(* IEC 61131-3 sources: Summary-ETFA22/ahorn/test/benchmark/dissertation/PPU/ST (part 7) *)

(* ---- Scenario8_Final_TODO.st ---- *)
FUNCTION_BLOCK Crane

    VAR_OUTPUT
        AnalogCranePressure : INT := INT#0;
        CraneLower : BOOL := FALSE;
        CraneTurnClockwise : BOOL := FALSE;
        CraneTurnCounterclockwise : BOOL := FALSE;
        MagazinVacuumOff : BOOL := FALSE;
        MagazinVacuumOn : BOOL := FALSE;
        StartCommandCrane : BOOL := FALSE;
    END_VAR

    VAR_INPUT
        CraneDown : BOOL := FALSE;
        CraneOnConveyor : BOOL := FALSE;
        CraneOnMagazin : BOOL := FALSE;
        CranePositionStamp : BOOL := FALSE;
        CraneSucked : BOOL := FALSE;
        CraneUp : BOOL := FALSE;
        MagazinCapacitiveSensor : BOOL := FALSE;
        MagazinOpticalSensor : BOOL := FALSE;
        SFCReset : BOOL := FALSE;
        SliderMovedOut : BOOL := FALSE;
        SliderNotMovedOut : BOOL := FALSE;
        StampLowered : BOOL := FALSE;
        StampSliderFilled : BOOL := FALSE;
        StampSliderSensorMovedOut : BOOL := FALSE;
        StartButtonMagazin : BOOL := FALSE;
        StartVar : BOOL := FALSE;
        WorkpieceReady : BOOL := FALSE;
    END_VAR

    VAR
        Duration1 : TIME := TIME#1500.0ms;
        SFCInit : BOOL := FALSE;
        TimeDelay_Timer : TON := (Q:=FALSE, PT:=UINT#0, IN:=FALSE, ET:=UINT#0);
        TimeDelay_Timer_Duration : TIME := TIME#50.0ms;
        TimeDelay_Timer_interconnect : BOOL := FALSE;
        Timer1 : TON := (Q:=FALSE, PT:=UINT#0, IN:=FALSE, ET:=UINT#0);
        actualtime1 : TIME := TIME#;
        interconnect : BOOL := FALSE;
        interconnectCraneStartCommand : BOOL := FALSE;
    END_VAR

    VAR
        SFCPause : BOOL := FALSE;
    END_VAR

    VAR
        __transit : BOOL := FALSE;
        _state : STATES_CRANE := STATES_CRANE#INIT;
    END_VAR

    ACTION Turn_Right_active
        CraneTurnClockwise := TRUE;
        CraneTurnCounterclockwise := FALSE;
    END_ACTION
    ACTION Crane_Turn_Left_White_active
        CraneTurnCounterclockwise := TRUE;
        CraneTurnClockwise := FALSE;
    END_ACTION
    ACTION Crane_Turn_Left_Metallic_active
        CraneTurnCounterclockwise := TRUE;
        CraneTurnClockwise := FALSE;
    END_ACTION
    ACTION Crane_Lift_Conveyor2_active
        CraneLower := FALSE;
    END_ACTION
    ACTION Crane_Turn_Right_From_Stamp_active
        CraneTurnClockwise := TRUE;
        CraneTurnCounterclockwise := FALSE;
    END_ACTION
    ACTION Suck_At_Stamp_active
        MagazinVacuumOn := TRUE;
        MagazinVacuumOff := FALSE;
    END_ACTION
    ACTION CraneTurnLeft_active
        CraneTurnCounterclockwise := TRUE;
        CraneTurnClockwise := FALSE;
    END_ACTION
    ACTION Crane_Turn_Left_From_Stamp_active
        CraneTurnClockwise := TRUE;
        CraneTurnCounterclockwise := FALSE;
    END_ACTION
    ACTION release_Black_active
        MagazinVacuumOn := FALSE;
        MagazinVacuumOff := TRUE;
    END_ACTION
    ACTION Crane_On_Stamp_Stop_Black_active
        CraneTurnClockwise := FALSE;
        CraneTurnCounterclockwise := FALSE;
    END_ACTION
    ACTION Reset_interconnect_active
        interconnect := FALSE;
        Timer1(IN := FALSE, PT := TIME#1ms);
    END_ACTION
    ACTION Crane_On_Stamp_White_active
        CraneTurnCounterclockwise := FALSE;
        CraneTurnClockwise := FALSE;
        CraneLower := TRUE;
    END_ACTION
    ACTION Crane_On_Stamp_Metallic_active
        CraneTurnCounterclockwise := FALSE;
        CraneTurnClockwise := FALSE;
        CraneLower := TRUE;
    END_ACTION
    ACTION Crane_Lift_Magazin_Metallic_active_0
        CraneLower := FALSE;
    END_ACTION
    ACTION TimeDelay_active
        TimeDelay_Timer(IN := TRUE, PT := TimeDelay_Timer_Duration);
        TimeDelay_Timer_interconnect := TimeDelay_Timer.Q;
    END_ACTION
    ACTION CraneLiftConveyor_active
        CraneLower := FALSE;
    END_ACTION
    ACTION Crane_Turn_Left_Back_To_Stamp_active
        CraneTurnCounterclockwise := TRUE;
        CraneTurnClockwise := FALSE;
    END_ACTION
    ACTION Crane_Init_2_active
        CraneLower := FALSE;
    END_ACTION
    ACTION Crane_Lower_active
        MagazinVacuumOn := TRUE;
        MagazinVacuumOff := FALSE;
        CraneLower := TRUE;
        AnalogCranePressure := INT#0;
    END_ACTION
    ACTION Crane_Lift_At_Stamp2_active
        CraneLower := FALSE;
    END_ACTION
    ACTION Crane_On_Stamp_Metallic2_active
        CraneTurnCounterclockwise := FALSE;
        CraneTurnClockwise := FALSE;
    END_ACTION
    ACTION CraneLiftMagazin_active
        CraneLower := FALSE;
    END_ACTION
    ACTION release_active
        MagazinVacuumOff := TRUE;
        MagazinVacuumOn := FALSE;
    END_ACTION
    ACTION Lower_Crane_active
        CraneLower := TRUE;
    END_ACTION
    ACTION Start_Crane_active
        CraneLower := FALSE;
        MagazinVacuumOff := TRUE;
        MagazinVacuumOn := FALSE;
        CraneTurnCounterclockwise := FALSE;
        CraneTurnClockwise := FALSE;
        StartVar := FALSE;
        StartCommandCrane := FALSE;
        IF (StartButtonMagazin = TRUE) THEN
            interconnectCraneStartCommand := TRUE;
        END_IF
    END_ACTION
    ACTION Crane_Go_Up_White_active
        CraneLower := FALSE;
    END_ACTION
    ACTION Crane_Init_active
        CraneLower := TRUE;
        interconnectCraneStartCommand := FALSE;
        AnalogCranePressure := INT#6000;
    END_ACTION
    ACTION Crane_Turn_Left_NOT_Metallic_Black_active
        CraneTurnCounterclockwise := TRUE;
        CraneTurnClockwise := FALSE;
    END_ACTION
    ACTION release_Workpiece_White_active
        MagazinVacuumOff := TRUE;
        MagazinVacuumOn := FALSE;
    END_ACTION
    ACTION Crane_On_Stamp_Metallic2_Lower_active
        CraneLower := TRUE;
    END_ACTION
    ACTION Crane_Turn_Left_Metallic2_active
        CraneTurnCounterclockwise := TRUE;
        CraneTurnClockwise := FALSE;
    END_ACTION
    ACTION Crane_Lift_NOT_Metallic_Black_active
        CraneLower := FALSE;
    END_ACTION
    ACTION Magazin_Stop_active
        CraneTurnClockwise := FALSE;
        CraneTurnCounterClockwise := FALSE;
    END_ACTION
    ACTION Crane_On_Conveyor_Not_Metallica_Black_active
        CraneTurnCounterclockwise := FALSE;
        CraneTurnClockwise := FALSE;
        CraneLower := TRUE;
    END_ACTION
    ACTION release_Workpiece_active
        MagazinVacuumOff := TRUE;
        MagazinVacuumOn := FALSE;
    END_ACTION
    ACTION No_Workpiece_ready_active_0
        MagazinVacuumOn := FALSE;
        MagazinVacuumOff := FALSE;
        CraneLower := FALSE;
    END_ACTION
    ACTION CraneOnConveyor_active
        CraneTurnCounterclockwise := FALSE;
        CraneTurnClockwise := FALSE;
        CraneLower := TRUE;
    END_ACTION
    ACTION Crane_Go_Up_active
        CraneLower := FALSE;
    END_ACTION
    ACTION Turn_Right_Final_active
        CraneTurnClockwise := TRUE;
        CraneTurnCounterclockwise := FALSE;
        AnalogCranePressure := INT#0;
    END_ACTION
    ACTION Suck_At_Stamp2_active
        MagazinVacuumOn := TRUE;
        MagazinVacuumOff := FALSE;
    END_ACTION
    ACTION Stamp_Pressure_Profile_Set_White_active
        AnalogCranePressure := INT#6000;
    END_ACTION
    ACTION Interstep_active
        StartCommandCrane := TRUE;
    END_ACTION
    ACTION Turn_Right_Black_active
        CraneTurnClockwise := TRUE;
        CraneTurnCounterclockwise := FALSE;
    END_ACTION
    ACTION Crane_On_Conveyor_Metallic2_active
        CraneTurnCounterclockwise := FALSE;
        CraneTurnClockwise := FALSE;
        CraneLower := TRUE;
    END_ACTION
    ACTION Crane_Lift_Conveyor_Black_active
        CraneLower := FALSE;
    END_ACTION
    ACTION Magazin_Stop_Final_active
        CraneTurnClockwise := FALSE;
        CraneTurnCounterClockwise := FALSE;
    END_ACTION
    ACTION Stamp_Pressure_Profile_Set_Metallic_active
        AnalogCranePressure := INT#7000;
    END_ACTION
    ACTION Crane_Lift_At_Stamp_active
        CraneLower := FALSE;
    END_ACTION
    ACTION Magazin_Stop_Black_active
        CraneTurnClockwise := FALSE;
        CraneTurnCounterclockwise := FALSE;
        MagazinVacuumOn := TRUE;
        MagazinVacuumOff := FALSE;
        CraneLower := TRUE;
    END_ACTION
    ACTION Crane_Lift_Magazin_White_active
        CraneLower := FALSE;
    END_ACTION
    ACTION pause_active
        Timer1(IN := CraneUP, PT := Duration1);
        interconnect := Timer1.Q;
    END_ACTION
    ACTION Crane_On_Conveyor_Metallic_active_0
        CraneTurnCounterclockwise := FALSE;
        CraneTurnClockwise := FALSE;
        CraneLower := TRUE;
    END_ACTION
    ACTION release2_active
        MagazinVacuumOff := TRUE;
        MagazinVacuumOn := FALSE;
    END_ACTION
    IF (SFCInit OR SFCReset) THEN
        AnalogCranePressure := INT#0;
        CraneDown := FALSE;
        CraneLower := FALSE;
        CraneOnConveyor := FALSE;
        CraneOnMagazin := FALSE;
        CranePositionStamp := FALSE;
        CraneSucked := FALSE;
        CraneTurnClockwise := FALSE;
        CraneTurnCounterclockwise := FALSE;
        CraneUp := FALSE;
        Duration1 := TIME#1500ms;
        MagazinCapacitiveSensor := FALSE;
        MagazinOpticalSensor := FALSE;
        MagazinVacuumOff := FALSE;
        MagazinVacuumOn := FALSE;
        SFCInit := FALSE;
        SFCReset := FALSE;
        SliderMovedOut := FALSE;
        SliderNotMovedOut := FALSE;
        StampLowered := FALSE;
        StampSliderFilled := FALSE;
        StampSliderSensorMovedOut := FALSE;
        StartButtonMagazin := FALSE;
        StartCommandCrane := FALSE;
        StartVar := FALSE;
        TimeDelay_Timer.ET := UINT#0;
        TimeDelay_Timer.IN := FALSE;
        TimeDelay_Timer.PT := UINT#0;
        TimeDelay_Timer.Q := FALSE;
        TimeDelay_Timer_Duration := TIME#50ms;
        TimeDelay_Timer_interconnect := FALSE;
        Timer1.ET := UINT#0;
        Timer1.IN := FALSE;
        Timer1.PT := UINT#0;
        Timer1.Q := FALSE;
        WorkpieceReady := FALSE;
        __transit := FALSE;
        _state := STATES_CRANE#INIT;
        actualtime1 := TIME#0ms;
        interconnect := FALSE;
        interconnectCraneStartCommand := FALSE;
    END_IF
    IF NOT (SFCInit OR SFCPause) THEN
        //Running pipeline step: edu.kit.iti.formal.automation.st.IntroduceStateEnumVariable

        //End of: edu.kit.iti.formal.automation.st.IntroduceStateEnumVariable

        //Running pipeline step: edu.kit.iti.formal.automation.st.TranslationSfcToStOld$IntroduceTransitVariable

        //End of: edu.kit.iti.formal.automation.st.TranslationSfcToStOld$IntroduceTransitVariable

        //Running pipeline step: edu.kit.iti.formal.automation.st.TranslationSfcToStOld$TheBigStateCase

        CASE _state OF
            STATES_CRANE#Init:
                __transit := FALSE;
                IF TRUE THEN
                    __transit := TRUE;
                    _state := STATES_CRANE#Start_Crane;
                END_IF

            STATES_CRANE#Start_Crane:
                __transit := FALSE;
                Start_Crane_active();
                IF interconnectCraneStartCommand THEN
                    __transit := TRUE;
                    _state := STATES_CRANE#Crane_Init;
                END_IF

            STATES_CRANE#Crane_Init:
                __transit := FALSE;
                Crane_Init_active();
                IF CraneDown THEN
                    __transit := TRUE;
                    _state := STATES_CRANE#Crane_Init_2;
                END_IF

            STATES_CRANE#Crane_Init_2:
                __transit := FALSE;
                Crane_Init_2_active();
                IF CraneUp THEN
                    __transit := TRUE;
                    _state := STATES_CRANE#Interstep;
                END_IF

            STATES_CRANE#Interstep:
                __transit := FALSE;
                Interstep_active();
                IF StartVar THEN
                    __transit := TRUE;
                    _state := STATES_CRANE#Interstep_2;
                END_IF

            STATES_CRANE#Interstep_2:
                __transit := FALSE;
                IF SliderMovedOut THEN
                    __transit := TRUE;
                    _state := STATES_CRANE#TimeDelay;
                END_IF

            STATES_CRANE#TimeDelay:
                __transit := FALSE;
                TimeDelay_active();
                IF TimeDelay_Timer_interconnect THEN
                    __transit := TRUE;
                    _state := STATES_CRANE#Interstep_3;
                END_IF

            STATES_CRANE#Interstep_3:
                __transit := FALSE;
                IF WorkpieceReady THEN
                    __transit := TRUE;
                    _state := STATES_CRANE#Turn_Right;
                ELSIF NOT WorkpieceReady THEN
                    __transit := TRUE;
                    _state := STATES_CRANE#No_Workpiece_ready;
                END_IF

            STATES_CRANE#Turn_Right:
                __transit := FALSE;
                Turn_Right_active();
                IF CraneOnMagazin THEN
                    __transit := TRUE;
                    _state := STATES_CRANE#Magazin_Stop;
                END_IF

            STATES_CRANE#Magazin_Stop:
                __transit := FALSE;
                Magazin_Stop_active();
                IF TRUE THEN
                    __transit := TRUE;
                    _state := STATES_CRANE#Crane_Lower;
                END_IF

            STATES_CRANE#Crane_Lower:
                __transit := FALSE;
                Crane_Lower_active();
                IF CraneSucked THEN
                    __transit := TRUE;
                    _state := STATES_CRANE#Step0;
                END_IF

            STATES_CRANE#Step0:
                __transit := FALSE;
                IF (NOT MagazinCapacitiveSensor AND NOT MagazinOpticalSensor) THEN
                    __transit := TRUE;
                    _state := STATES_CRANE#Crane_Lift_Magazin;
                ELSIF (MagazinCapacitiveSensor AND MagazinOpticalSensor) THEN
                    __transit := TRUE;
                    _state := STATES_CRANE#Stamp_Pressure_Profile_Set_Metallic;
                ELSIF (NOT MagazinCapacitiveSensor AND MagazinOpticalSensor) THEN
                    __transit := TRUE;
                    _state := STATES_CRANE#Stamp_Pressure_Profile_Set_White;
                ELSIF (MagazinCapacitiveSensor AND MagazinOpticalSensor) THEN
                    __transit := TRUE;
                    _state := STATES_CRANE#Stamp_Pressure_Profile_Set_Metallic;
                ELSIF (NOT MagazinCapacitiveSensor AND MagazinOpticalSensor) THEN
                    __transit := TRUE;
                    _state := STATES_CRANE#Stamp_Pressure_Profile_Set_White;
                END_IF

            STATES_CRANE#Crane_Lift_Magazin:
                __transit := FALSE;
                CraneLiftMagazin_active();
                IF CraneUp THEN
                    __transit := TRUE;
                    _state := STATES_CRANE#Crane_Turn_Left_NOT_Metallic;
                END_IF

            STATES_CRANE#Crane_Turn_Left_NOT_Metallic:
                __transit := FALSE;
                CraneTurnLeft_active();
                IF CraneOnConveyor THEN
                    __transit := TRUE;
                    _state := STATES_CRANE#Crane_On_Conveyor;
                END_IF

            STATES_CRANE#Crane_On_Conveyor:
                __transit := FALSE;
                CraneOnConveyor_active();
                IF CraneDown THEN
                    __transit := TRUE;
                    _state := STATES_CRANE#release;
                END_IF

            STATES_CRANE#Stamp_Pressure_Profile_Set_Metallic:
                __transit := FALSE;
                Stamp_Pressure_Profile_Set_Metallic_active();
                IF TRUE THEN
                    __transit := TRUE;
                    _state := STATES_CRANE#Crane_Lift_Magazin_Metallic;
                END_IF

            STATES_CRANE#Crane_Lift_Magazin_Metallic:
                __transit := FALSE;
                Crane_Lift_Magazin_Metallic_active_0();
                IF CraneUp THEN
                    __transit := TRUE;
                    _state := STATES_CRANE#Crane_Turn_Left_Metallic;
                END_IF

            STATES_CRANE#Crane_Turn_Left_Metallic:
                __transit := FALSE;
                Crane_Turn_Left_Metallic_active();
                IF CranePositionStamp THEN
                    __transit := TRUE;
                    _state := STATES_CRANE#Crane_On_Stamp_Metallic;
                END_IF

            STATES_CRANE#Crane_On_Stamp_Metallic:
                __transit := FALSE;
                Crane_On_Stamp_Metallic_active();
                IF CraneDown THEN
                    __transit := TRUE;
                    _state := STATES_CRANE#release_Workpiece;
                END_IF

            STATES_CRANE#release_Workpiece:
                __transit := FALSE;
                release_Workpiece_active();
                IF TRUE THEN
                    __transit := TRUE;
                    _state := STATES_CRANE#Crane_Go_Up;
                END_IF

            STATES_CRANE#Crane_Go_Up:
                __transit := FALSE;
                Crane_Go_Up_active();
                IF CraneUp THEN
                    __transit := TRUE;
                    _state := STATES_CRANE#Step3;
                END_IF

            STATES_CRANE#Stamp_Pressure_Profile_Set_White:
                __transit := FALSE;
                Stamp_Pressure_Profile_Set_White_active();
                IF TRUE THEN
                    __transit := TRUE;
                    _state := STATES_CRANE#Crane_Lift_Magazine_White;
                END_IF

            STATES_CRANE#Crane_Lift_Magazine_White:
                __transit := FALSE;
                Crane_Lift_Magazin_White_active();
                IF CraneUp THEN
                    __transit := TRUE;
                    _state := STATES_CRANE#Crane_Turn_Left_White;
                END_IF

            STATES_CRANE#Crane_Turn_Left_White:
                __transit := FALSE;
                Crane_Turn_Left_White_active();
                IF CranePositionStamp THEN
                    __transit := TRUE;
                    _state := STATES_CRANE#Crane_On_Stamp_White;
                END_IF

            STATES_CRANE#Crane_On_Stamp_White:
                __transit := FALSE;
                Crane_On_Stamp_White_active();
                IF CraneDown THEN
                    __transit := TRUE;
                    _state := STATES_CRANE#release_Workpiece_White;
                END_IF

            STATES_CRANE#release_Workpiece_White:
                __transit := FALSE;
                release_Workpiece_White_active();
                IF TRUE THEN
                    __transit := TRUE;
                    _state := STATES_CRANE#Crane_Go_Up_White;
                END_IF

            STATES_CRANE#Crane_Go_Up_White:
                __transit := FALSE;
                Crane_Go_Up_White_active();
                IF CraneUp THEN
                    __transit := TRUE;
                    _state := STATES_CRANE#Step3;
                END_IF

            STATES_CRANE#Step3:
                __transit := FALSE;
                IF WorkpieceReady THEN
                    __transit := TRUE;
                    _state := STATES_CRANE#Step2;
                ELSIF NOT WorkpieceReady THEN
                    __transit := TRUE;
                    _state := STATES_CRANE#Step4;
                END_IF

            STATES_CRANE#Step2:
                __transit := FALSE;
                IF (MagazinCapacitiveSensor OR MagazinOpticalSensor) THEN
                    __transit := TRUE;
                    _state := STATES_CRANE#pause;
                ELSIF (NOT MagazinCapacitiveSensor AND NOT MagazinOpticalSensor) THEN
                    __transit := TRUE;
                    _state := STATES_CRANE#Turn_Right_Black;
                END_IF

            STATES_CRANE#pause:
                __transit := FALSE;
                pause_active();
                IF interconnect THEN
                    __transit := TRUE;
                    _state := STATES_CRANE#Reset_interconnect;
                ELSIF interconnect THEN
                    __transit := TRUE;
                    _state := STATES_CRANE#Reset_interconnect;
                END_IF

            STATES_CRANE#Turn_Right_Black:
                __transit := FALSE;
                Turn_Right_Black_active();
                IF CraneOnMagazin THEN
                    __transit := TRUE;
                    _state := STATES_CRANE#Magazin_Stop_Black;
                END_IF

            STATES_CRANE#Magazin_Stop_Black:
                __transit := FALSE;
                Magazin_Stop_Black_active();
                IF CraneSucked THEN
                    __transit := TRUE;
                    _state := STATES_CRANE#Crane_Lift_NOT_Metallic_Black;
                END_IF

            STATES_CRANE#Crane_Lift_NOT_Metallic_Black:
                __transit := FALSE;
                Crane_Lift_NOT_Metallic_Black_active();
                IF CraneUp THEN
                    __transit := TRUE;
                    _state := STATES_CRANE#Crane_Turn_Left_NOT_Metallic_Black;
                END_IF

            STATES_CRANE#Crane_Turn_Left_NOT_Metallic_Black:
                __transit := FALSE;
                Crane_Turn_Left_NOT_Metallic_Black_active();
                IF CraneOnConveyor THEN
                    __transit := TRUE;
                    _state := STATES_CRANE#Crane_On_Conveyor_Not_Metallica_Black;
                END_IF

            STATES_CRANE#Crane_On_Conveyor_Not_Metallica_Black:
                __transit := FALSE;
                Crane_On_Conveyor_Not_Metallica_Black_active();
                IF CraneDown THEN
                    __transit := TRUE;
                    _state := STATES_CRANE#release_Black;
                END_IF

            STATES_CRANE#release_Black:
                __transit := FALSE;
                release_Black_active();
                IF TRUE THEN
                    __transit := TRUE;
                    _state := STATES_CRANE#Crane_Lift_Conveyor_Black;
                END_IF

            STATES_CRANE#Crane_Lift_Conveyor_Black:
                __transit := FALSE;
                Crane_Lift_Conveyor_Black_active();
                IF CraneUp THEN
                    __transit := TRUE;
                    _state := STATES_CRANE#Crane_Turn_Left_Back_To_Stamp;
                END_IF

            STATES_CRANE#Crane_Turn_Left_Back_To_Stamp:
                __transit := FALSE;
                Crane_Turn_Left_Back_To_Stamp_active();
                IF CranePositionStamp THEN
                    __transit := TRUE;
                    _state := STATES_CRANE#Crane_On_Stamp_Stop_Black;
                END_IF

            STATES_CRANE#Crane_On_Stamp_Stop_Black:
                __transit := FALSE;
                Crane_On_Stamp_Stop_Black_active();
                IF TRUE THEN
                    __transit := TRUE;
                    _state := STATES_CRANE#Reset_interconnect;
                ELSIF TRUE THEN
                    __transit := TRUE;
                    _state := STATES_CRANE#Reset_interconnect;
                END_IF

            STATES_CRANE#Step4:
                __transit := FALSE;
                IF TRUE THEN
                    __transit := TRUE;
                    _state := STATES_CRANE#Interstep;
                END_IF

            STATES_CRANE#Reset_interconnect:
                __transit := FALSE;
                Reset_interconnect_active();
                IF SliderMovedOut THEN
                    __transit := TRUE;
                    _state := STATES_CRANE#Lower_Crane;
                END_IF

            STATES_CRANE#Lower_Crane:
                __transit := FALSE;
                Lower_Crane_active();
                IF CraneDown THEN
                    __transit := TRUE;
                    _state := STATES_CRANE#Suck_At_Stamp;
                END_IF

            STATES_CRANE#Suck_At_Stamp:
                __transit := FALSE;
                Suck_At_Stamp_active();
                IF CraneSucked THEN
                    __transit := TRUE;
                    _state := STATES_CRANE#Crane_Lift_At_Stamp;
                END_IF

            STATES_CRANE#Crane_Lift_At_Stamp:
                __transit := FALSE;
                Crane_Lift_At_Stamp_active();
                IF CraneUp THEN
                    __transit := TRUE;
                    _state := STATES_CRANE#Crane_Turn_Left_From_Stamp;
                END_IF

            STATES_CRANE#Crane_Turn_Left_From_Stamp:
                __transit := FALSE;
                Crane_Turn_Left_From_Stamp_active();
                IF CraneOnConveyor THEN
                    __transit := TRUE;
                    _state := STATES_CRANE#Crane_On_Conveyor_Metallic;
                END_IF

            STATES_CRANE#Crane_On_Conveyor_Metallic:
                __transit := FALSE;
                Crane_On_Conveyor_Metallic_active_0();
                IF CraneDown THEN
                    __transit := TRUE;
                    _state := STATES_CRANE#release;
                END_IF

            STATES_CRANE#release:
                __transit := FALSE;
                release_active();
                IF TRUE THEN
                    __transit := TRUE;
                    _state := STATES_CRANE#Crane_Lift_Conveyor;
                END_IF

            STATES_CRANE#Crane_Lift_Conveyor:
                __transit := FALSE;
                CraneLiftConveyor_active();
                IF TRUE THEN
                    __transit := TRUE;
                    _state := STATES_CRANE#Interstep;
                END_IF

            STATES_CRANE#No_Workpiece_ready:
                __transit := FALSE;
                No_Workpiece_ready_active_0();
                IF StampSliderFilled THEN
                    __transit := TRUE;
                    _state := STATES_CRANE#Crane_Turn_Left_Metallic2;
                ELSIF NOT StampSliderFilled THEN
                    __transit := TRUE;
                    _state := STATES_CRANE#Turn_Right_Final;
                END_IF

            STATES_CRANE#Crane_Turn_Left_Metallic2:
                __transit := FALSE;
                Crane_Turn_Left_Metallic2_active();
                IF CranePositionStamp THEN
                    __transit := TRUE;
                    _state := STATES_CRANE#Crane_On_Stamp_Metallic2;
                END_IF

            STATES_CRANE#Crane_On_Stamp_Metallic2:
                __transit := FALSE;
                Crane_On_Stamp_Metallic2_active();
                IF StampLowered THEN
                    __transit := TRUE;
                    _state := STATES_CRANE#Interstep_4;
                END_IF

            STATES_CRANE#Interstep_4:
                __transit := FALSE;
                IF StampSliderSensorMovedOut THEN
                    __transit := TRUE;
                    _state := STATES_CRANE#Crane_On_Stamp_Metallic2_Lower;
                END_IF

            STATES_CRANE#Crane_On_Stamp_Metallic2_Lower:
                __transit := FALSE;
                Crane_On_Stamp_Metallic2_Lower_active();
                IF CraneDown THEN
                    __transit := TRUE;
                    _state := STATES_CRANE#Suck_At_Stamp2;
                END_IF

            STATES_CRANE#Suck_At_Stamp2:
                __transit := FALSE;
                Suck_At_Stamp2_active();
                IF CraneSucked THEN
                    __transit := TRUE;
                    _state := STATES_CRANE#Crane_Lift_At_Stamp2;
                END_IF

            STATES_CRANE#Crane_Lift_At_Stamp2:
                __transit := FALSE;
                Crane_Lift_At_Stamp2_active();
                IF CraneUp THEN
                    __transit := TRUE;
                    _state := STATES_CRANE#Crane_Turn_Right_From_Stamp;
                END_IF

            STATES_CRANE#Crane_Turn_Right_From_Stamp:
                __transit := FALSE;
                Crane_Turn_Right_From_Stamp_active();
                IF CraneOnConveyor THEN
                    __transit := TRUE;
                    _state := STATES_CRANE#Crane_On_Conveyor_Metallic2;
                END_IF

            STATES_CRANE#Crane_On_Conveyor_Metallic2:
                __transit := FALSE;
                Crane_On_Conveyor_Metallic2_active();
                IF CraneDown THEN
                    __transit := TRUE;
                    _state := STATES_CRANE#release2;
                END_IF

            STATES_CRANE#release2:
                __transit := FALSE;
                release2_active();
                IF TRUE THEN
                    __transit := TRUE;
                    _state := STATES_CRANE#Crane_Lift_Conveyor2;
                END_IF

            STATES_CRANE#Crane_Lift_Conveyor2:
                __transit := FALSE;
                Crane_Lift_Conveyor2_active();
                IF TRUE THEN
                    __transit := TRUE;
                    _state := STATES_CRANE#Interstep;
                ELSIF TRUE THEN
                    __transit := TRUE;
                    _state := STATES_CRANE#Interstep;
                END_IF

            STATES_CRANE#Turn_Right_Final:
                __transit := FALSE;
                Turn_Right_Final_active();
                IF CraneOnMagazin THEN
                    __transit := TRUE;
                    _state := STATES_CRANE#Magazin_Stop_Final;
                END_IF

            STATES_CRANE#Magazin_Stop_Final:
                __transit := FALSE;
                Magazin_Stop_Final_active();
                IF TRUE THEN
                    __transit := TRUE;
                    _state := STATES_CRANE#Start_Crane;
                END_IF

                    END_CASE
        //End of: edu.kit.iti.formal.automation.st.TranslationSfcToStOld$TheBigStateCase

        //Running pipeline step: edu.kit.iti.formal.automation.st.SfcFlagIntroduction

    END_IF
    //End of: edu.kit.iti.formal.automation.st.SfcFlagIntroduction

END_FUNCTION_BLOCK

FUNCTION_BLOCK Magazin

    VAR_INPUT
        CraneDown : BOOL := FALSE;
        CraneOnConveyor : BOOL := FALSE;
        CraneOnMagazin : BOOL := FALSE;
        CraneSucked : BOOL := FALSE;
        CraneUp : BOOL := FALSE;
        SFCReset : BOOL := FALSE;
        SliderMovedOut : BOOL := FALSE;
        SliderNotMovedOut : BOOL := FALSE;
        StartButtonMagazin : BOOL := FALSE;
        StartVar : BOOL := FALSE;
        WorkpieceReady : BOOL := FALSE;
    END_VAR

    VAR_OUTPUT
        CraneLower : BOOL := FALSE;
        CraneTurnClockwise : BOOL := FALSE;
        CraneTurnCounterclockwise : BOOL := FALSE;
        MagazinGreenLamp : BOOL := FALSE;
        MagazinSlider : BOOL := FALSE;
        MagazinVacuumOff : BOOL := FALSE;
        MagazinVacuumOn : BOOL := FALSE;
        MagazinWhiteLamp : BOOL := FALSE;
        StartCommandMagazin : BOOL := FALSE;
    END_VAR

    VAR
        SFCInit : BOOL := FALSE;
        interconnectMagazinStartCommand : BOOL := FALSE;
    END_VAR

    VAR
        SFCPause : BOOL := FALSE;
    END_VAR

    VAR
        __transit : BOOL := FALSE;
        _state : STATES_MAGAZIN := STATES_MAGAZIN#INIT;
    END_VAR

    ACTION Magazin_Init_2_active
        MagazinSlider := FALSE;
    END_ACTION
    ACTION Start_Magazin_active
        MagazinSlider := FALSE;
        MagazinGreenLamp := FALSE;
        StartVar := FALSE;
        StartCommandMagazin := FALSE;
        IF (StartButtonMagazin = TRUE) THEN
            interconnectMagazinStartCommand := TRUE;
        END_IF
    END_ACTION
    ACTION Green_Lamp_active
        MagazinGreenLamp := TRUE;
        interconnectMagazinStartCommand := FALSE;
    END_ACTION
    ACTION SliderMoveBack_active
        IF ((SliderMovedOut = TRUE) AND (SliderNotMovedOut = FALSE)) THEN
            MagazinSlider := FALSE;
        END_IF
    END_ACTION
    ACTION convey_active
        IF SliderNotMovedOut THEN
            MagazinSlider := TRUE;
        END_IF
    END_ACTION
    ACTION Magazin_Init_active
        MagazinSlider := TRUE;
    END_ACTION
    ACTION Interstep_active
        StartCommandMagazin := TRUE;
    END_ACTION
    IF (SFCInit OR SFCReset) THEN
        CraneDown := FALSE;
        CraneLower := FALSE;
        CraneOnConveyor := FALSE;
        CraneOnMagazin := FALSE;
        CraneSucked := FALSE;
        CraneTurnClockwise := FALSE;
        CraneTurnCounterclockwise := FALSE;
        CraneUp := FALSE;
        MagazinGreenLamp := FALSE;
        MagazinSlider := FALSE;
        MagazinVacuumOff := FALSE;
        MagazinVacuumOn := FALSE;
        MagazinWhiteLamp := FALSE;
        SFCInit := FALSE;
        SFCReset := FALSE;
        SliderMovedOut := FALSE;
        SliderNotMovedOut := FALSE;
        StartButtonMagazin := FALSE;
        StartCommandMagazin := FALSE;
        StartVar := FALSE;
        WorkpieceReady := FALSE;
        __transit := FALSE;
        _state := STATES_MAGAZIN#INIT;
        interconnectMagazinStartCommand := FALSE;
    END_IF
    IF NOT (SFCInit OR SFCPause) THEN
        //Running pipeline step: edu.kit.iti.formal.automation.st.IntroduceStateEnumVariable

        //End of: edu.kit.iti.formal.automation.st.IntroduceStateEnumVariable

        //Running pipeline step: edu.kit.iti.formal.automation.st.TranslationSfcToStOld$IntroduceTransitVariable

        //End of: edu.kit.iti.formal.automation.st.TranslationSfcToStOld$IntroduceTransitVariable

        //Running pipeline step: edu.kit.iti.formal.automation.st.TranslationSfcToStOld$TheBigStateCase

        CASE _state OF
            STATES_MAGAZIN#Init:
                __transit := FALSE;
                IF TRUE THEN
                    __transit := TRUE;
                    _state := STATES_MAGAZIN#Start_Magazin;
                END_IF

            STATES_MAGAZIN#Start_Magazin:
                __transit := FALSE;
                Start_Magazin_active();
                IF interconnectMagazinStartCommand THEN
                    __transit := TRUE;
                    _state := STATES_MAGAZIN#Green_Lamp;
                END_IF

            STATES_MAGAZIN#Green_Lamp:
                __transit := FALSE;
                Green_Lamp_active();
                IF TRUE THEN
                    __transit := TRUE;
                    _state := STATES_MAGAZIN#Magazin_Init;
                END_IF

            STATES_MAGAZIN#Magazin_Init:
                __transit := FALSE;
                Magazin_Init_active();
                IF TRUE THEN
                    __transit := TRUE;
                    _state := STATES_MAGAZIN#Magazin_Init_2;
                END_IF

            STATES_MAGAZIN#Magazin_Init_2:
                __transit := FALSE;
                Magazin_Init_2_active();
                IF TRUE THEN
                    __transit := TRUE;
                    _state := STATES_MAGAZIN#Interstep;
                END_IF

            STATES_MAGAZIN#Interstep:
                __transit := FALSE;
                Interstep_active();
                IF StartVar THEN
                    __transit := TRUE;
                    _state := STATES_MAGAZIN#convey;
                END_IF

            STATES_MAGAZIN#convey:
                __transit := FALSE;
                convey_active();
                IF CraneOnMagazin THEN
                    __transit := TRUE;
                    _state := STATES_MAGAZIN#Step0;
                END_IF

            STATES_MAGAZIN#Step0:
                __transit := FALSE;
                IF CraneDown THEN
                    __transit := TRUE;
                    _state := STATES_MAGAZIN#Slider_Move_Back;
                END_IF

            STATES_MAGAZIN#Slider_Move_Back:
                __transit := FALSE;
                SliderMoveBack_active();
                IF CraneUp THEN
                    __transit := TRUE;
                    _state := STATES_MAGAZIN#Step1;
                END_IF

            STATES_MAGAZIN#Step1:
                __transit := FALSE;
                IF CraneOnConveyor THEN
                    __transit := TRUE;
                    _state := STATES_MAGAZIN#Interstep;
                END_IF

                    END_CASE
        //End of: edu.kit.iti.formal.automation.st.TranslationSfcToStOld$TheBigStateCase

        //Running pipeline step: edu.kit.iti.formal.automation.st.SfcFlagIntroduction

    END_IF
    //End of: edu.kit.iti.formal.automation.st.SfcFlagIntroduction

END_FUNCTION_BLOCK

FUNCTION_BLOCK Stamp

    VAR_INPUT
        CraneDown : BOOL := FALSE;
        CraneOnConveyor : BOOL := FALSE;
        CranePositionStamp : BOOL := FALSE;
        CraneSucked : BOOL := FALSE;
        CraneUp : BOOL := FALSE;
        SFCReset : BOOL := FALSE;
        StampLowered : BOOL := FALSE;
        StampSliderFilled : BOOL := FALSE;
        StampSliderSensorMovedIn : BOOL := FALSE;
        StampSliderSensorMovedOut : BOOL := FALSE;
        StampStartButton : BOOL := FALSE;
        StampUp : BOOL := FALSE;
        StartVar : BOOL := FALSE;
    END_VAR

    VAR
        Duration : TIME := TIME#500.0ms;
        SFCInit : BOOL := FALSE;
        Timer : TON := (Q:=FALSE, PT:=UINT#0, IN:=FALSE, ET:=UINT#0);
        interconnect : BOOL := FALSE;
        interconnectStampStartCommand : BOOL := FALSE;
    END_VAR

    VAR
        SFCPause : BOOL := FALSE;
    END_VAR

    VAR_OUTPUT
        StampGreenLamp : BOOL := FALSE;
        StampPressure : BOOL := FALSE;
        StampPusher : BOOL := FALSE;
        StampSliderMovedIn : BOOL := FALSE;
        StampSliderMovedOut : BOOL := FALSE;
        StampWhiteLamp : BOOL := FALSE;
        StartCommandStamp : BOOL := FALSE;
    END_VAR

    VAR
        __transit : BOOL := FALSE;
        _state : STATES_STAMP := STATES_STAMP#INIT;
    END_VAR

    ACTION StampSliderForward_active
        StampPusher := FALSE;
        StampSliderMovedOut := TRUE;
        IF ((StampLowered = FALSE) AND (StampUp = TRUE)) THEN
            interconnect := FALSE;
        END_IF
        Timer(IN := FALSE, PT := TIME#1ms);
    END_ACTION
    ACTION Start_Stamp_active
        StampSliderMovedOut := FALSE;
        StampSliderMovedIn := FALSE;
        StampPusher := FALSE;
        StampGreenLamp := FALSE;
        StampPressure := FALSE;
        StartCommandStamp := FALSE;
        IF (StampStartButton = TRUE) THEN
            interconnectStampStartCommand := TRUE;
        END_IF
    END_ACTION
    ACTION Step1_active
        Timer(IN := StampLowered, PT := TIME#0ms);
        interconnect := Timer.Q;
    END_ACTION
    ACTION Green_Lamp_active
        StampGreenLamp := TRUE;
        interconnectStampStartCommand := FALSE;
    END_ACTION
    ACTION Stamp_Init_4_active
        StampPusher := FALSE;
    END_ACTION
    ACTION Interstep_active
        StartCommandStamp := TRUE;
    END_ACTION
    ACTION Stamp_Init_2_active
        StampSliderMovedIn := FALSE;
        StampSliderMovedOut := TRUE;
    END_ACTION
    ACTION Stamp_Init_3_active
        StampPusher := TRUE;
    END_ACTION
    ACTION Stamp_Init_1_active
        StampSliderMovedIn := TRUE;
        StampSliderMovedOut := FALSE;
    END_ACTION
    ACTION StampProcess_active
        StampSliderMovedIn := FALSE;
        StampPusher := TRUE;
    END_ACTION
    ACTION StampSliderBack_active
        StampSliderMovedIn := TRUE;
        StampSliderMovedOut := FALSE;
    END_ACTION
    IF (SFCInit OR SFCReset) THEN
        CraneDown := FALSE;
        CraneOnConveyor := FALSE;
        CranePositionStamp := FALSE;
        CraneSucked := FALSE;
        CraneUp := FALSE;
        Duration := TIME#500ms;
        SFCInit := FALSE;
        SFCReset := FALSE;
        StampGreenLamp := FALSE;
        StampLowered := FALSE;
        StampPressure := FALSE;
        StampPusher := FALSE;
        StampSliderFilled := FALSE;
        StampSliderMovedIn := FALSE;
        StampSliderMovedOut := FALSE;
        StampSliderSensorMovedIn := FALSE;
        StampSliderSensorMovedOut := FALSE;
        StampStartButton := FALSE;
        StampUp := FALSE;
        StampWhiteLamp := FALSE;
        StartCommandStamp := FALSE;
        StartVar := FALSE;
        Timer.ET := UINT#0;
        Timer.IN := FALSE;
        Timer.PT := UINT#0;
        Timer.Q := FALSE;
        __transit := FALSE;
        _state := STATES_STAMP#INIT;
        interconnect := FALSE;
        interconnectStampStartCommand := FALSE;
    END_IF
    IF NOT (SFCInit OR SFCPause) THEN
        //Running pipeline step: edu.kit.iti.formal.automation.st.IntroduceStateEnumVariable

        //End of: edu.kit.iti.formal.automation.st.IntroduceStateEnumVariable

        //Running pipeline step: edu.kit.iti.formal.automation.st.TranslationSfcToStOld$IntroduceTransitVariable

        //End of: edu.kit.iti.formal.automation.st.TranslationSfcToStOld$IntroduceTransitVariable

        //Running pipeline step: edu.kit.iti.formal.automation.st.TranslationSfcToStOld$TheBigStateCase

        CASE _state OF
            STATES_STAMP#Init:
                __transit := FALSE;
                IF TRUE THEN
                    __transit := TRUE;
                    _state := STATES_STAMP#Start_Stamp;
                END_IF

            STATES_STAMP#Start_Stamp:
                __transit := FALSE;
                Start_Stamp_active();
                IF interconnectStampStartCommand THEN
                    __transit := TRUE;
                    _state := STATES_STAMP#Green_Lamp;
                END_IF

            STATES_STAMP#Green_Lamp:
                __transit := FALSE;
                Green_Lamp_active();
                IF TRUE THEN
                    __transit := TRUE;
                    _state := STATES_STAMP#Stamp_Init_1;
                END_IF

            STATES_STAMP#Stamp_Init_1:
                __transit := FALSE;
                Stamp_Init_1_active();
                IF StampSliderSensorMovedIn THEN
                    __transit := TRUE;
                    _state := STATES_STAMP#Stamp_Init_2;
                END_IF

            STATES_STAMP#Stamp_Init_2:
                __transit := FALSE;
                Stamp_Init_2_active();
                IF StampSliderSensorMovedOut THEN
                    __transit := TRUE;
                    _state := STATES_STAMP#Stamp_Init_3;
                END_IF

            STATES_STAMP#Stamp_Init_3:
                __transit := FALSE;
                Stamp_Init_3_active();
                IF StampLowered THEN
                    __transit := TRUE;
                    _state := STATES_STAMP#Stamp_Init_4;
                END_IF

            STATES_STAMP#Stamp_Init_4:
                __transit := FALSE;
                Stamp_Init_4_active();
                IF StampUp THEN
                    __transit := TRUE;
                    _state := STATES_STAMP#Interstep;
                END_IF

            STATES_STAMP#Interstep:
                __transit := FALSE;
                Interstep_active();
                IF StartVar THEN
                    __transit := TRUE;
                    _state := STATES_STAMP#Interstep_2;
                END_IF

            STATES_STAMP#Interstep_2:
                __transit := FALSE;
                IF StampSliderFilled THEN
                    __transit := TRUE;
                    _state := STATES_STAMP#Step0;
                END_IF

            STATES_STAMP#Step0:
                __transit := FALSE;
                IF CraneUp THEN
                    __transit := TRUE;
                    _state := STATES_STAMP#StampSliderBack;
                END_IF

            STATES_STAMP#StampSliderBack:
                __transit := FALSE;
                StampSliderBack_active();
                IF StampSliderSensorMovedIn THEN
                    __transit := TRUE;
                    _state := STATES_STAMP#StampProcess;
                END_IF

            STATES_STAMP#StampProcess:
                __transit := FALSE;
                StampProcess_active();
                IF StampLowered THEN
                    __transit := TRUE;
                    _state := STATES_STAMP#Step1;
                END_IF

            STATES_STAMP#Step1:
                __transit := FALSE;
                Step1_active();
                IF interconnect THEN
                    __transit := TRUE;
                    _state := STATES_STAMP#StampSliderForward;
                END_IF

            STATES_STAMP#StampSliderForward:
                __transit := FALSE;
                StampSliderForward_active();
                IF StampSliderMovedOut THEN
                    __transit := TRUE;
                    _state := STATES_STAMP#Step2;
                END_IF

            STATES_STAMP#Step2:
                __transit := FALSE;
                IF (CraneOnConveyor AND NOT StampSliderFilled) THEN
                    __transit := TRUE;
                    _state := STATES_STAMP#Interstep;
                END_IF

                    END_CASE
        //End of: edu.kit.iti.formal.automation.st.TranslationSfcToStOld$TheBigStateCase

        //Running pipeline step: edu.kit.iti.formal.automation.st.SfcFlagIntroduction

    END_IF
    //End of: edu.kit.iti.formal.automation.st.SfcFlagIntroduction

END_FUNCTION_BLOCK

PROGRAM Main
    VAR_OUTPUT
        Actuator_AnalogCranePressure : INT := INT#0;
        Actuator_CraneLower : BOOL := FALSE;
        Actuator_CraneTurnClockwise : BOOL := FALSE;
        Actuator_CraneTurnCounterclockwise : BOOL := FALSE;
        Actuator_MagazinGreenLamp : BOOL := FALSE;
        Actuator_MagazinSlider : BOOL := FALSE;
        Actuator_MagazinVacuumOff : BOOL := FALSE;
        Actuator_MagazinVacuumOn : BOOL := FALSE;
        Actuator_MagazinWhiteLamp : BOOL := FALSE;
        Actuator_StampGreenLamp : BOOL := FALSE;
        Actuator_StampPusher : BOOL := FALSE;
        Actuator_StampSliderMovedIn : BOOL := FALSE;
        Actuator_StampSliderMovedOut : BOOL := FALSE;
        Actuator_StampWhiteLamp : BOOL := FALSE;
    END_VAR

    VAR
        Crane : Crane := (SliderMovedOut:=FALSE, CraneTurnCounterclockwise:=FALSE, WorkpieceReady:=FALSE, StampLowered:=FALSE, Duration1:=TIME#1500.0ms, StampSliderSensorMovedOut:=FALSE, TimeDelay_Timer_interconnect:=FALSE, CraneOnConveyor:=FALSE, MagazinOpticalSensor:=FALSE, CranePositionStamp:=FALSE, StartVar:=FALSE, StartButtonMagazin:=FALSE, CraneOnMagazin:=FALSE, actualtime1:=TIME#, AnalogCranePressure:=INT#0, SFCReset:=FALSE, MagazinVacuumOff:=FALSE, CraneSucked:=FALSE, MagazinVacuumOn:=FALSE, interconnectCraneStartCommand:=FALSE, SFCInit:=FALSE, StartCommandCrane:=FALSE, TimeDelay_Timer_Duration:=TIME#50.0ms, interconnect:=FALSE, StampSliderFilled:=FALSE, CraneTurnClockwise:=FALSE, CraneUp:=FALSE, MagazinCapacitiveSensor:=FALSE, CraneLower:=FALSE, SliderNotMovedOut:=FALSE, CraneDown:=FALSE, TimeDelay_Timer:=(Q:=FALSE, PT:=UINT#0, IN:=FALSE, ET:=UINT#0), Timer1:=(Q:=FALSE, PT:=UINT#0, IN:=FALSE, ET:=UINT#0));
        Mag : Magazin := (SliderMovedOut:=FALSE, MagazinGreenLamp:=FALSE, interconnectMagazinStartCommand:=FALSE, SFCReset:=FALSE, CraneTurnCounterclockwise:=FALSE, MagazinVacuumOff:=FALSE, WorkpieceReady:=FALSE, CraneSucked:=FALSE, MagazinSlider:=FALSE, MagazinVacuumOn:=FALSE, MagazinWhiteLamp:=FALSE, SFCInit:=FALSE, StartCommandMagazin:=FALSE, CraneOnConveyor:=FALSE, CraneTurnClockwise:=FALSE, CraneUp:=FALSE, StartVar:=FALSE, CraneLower:=FALSE, SliderNotMovedOut:=FALSE, StartButtonMagazin:=FALSE, CraneOnMagazin:=FALSE, CraneDown:=FALSE);
        Stamp : Stamp := (StampLowered:=FALSE, StampSliderSensorMovedOut:=FALSE, interconnectStampStartCommand:=FALSE, CraneOnConveyor:=FALSE, CranePositionStamp:=FALSE, StampSliderMovedOut:=FALSE, StartVar:=FALSE, StampPusher:=FALSE, StampWhiteLamp:=FALSE, StampPressure:=FALSE, SFCReset:=FALSE, StampGreenLamp:=FALSE, CraneSucked:=FALSE, Duration:=TIME#500.0ms, SFCInit:=FALSE, StampStartButton:=FALSE, StampSliderSensorMovedIn:=FALSE, interconnect:=FALSE, StampSliderFilled:=FALSE, CraneUp:=FALSE, StampSliderMovedIn:=FALSE, Timer:=(Q:=FALSE, PT:=UINT#0, IN:=FALSE, ET:=UINT#0), StartCommandStamp:=FALSE, CraneDown:=FALSE, StampUp:=FALSE);
    END_VAR

    VAR_INPUT
        Sensor_CraneDown : BOOL := FALSE;
        Sensor_CraneOnConveyor : BOOL := FALSE;
        Sensor_CraneOnMagazin : BOOL := FALSE;
        Sensor_CranePosition : BOOL := FALSE;
        Sensor_CranePositionStamp : BOOL := FALSE;
        Sensor_CraneSucked : BOOL := FALSE;
        Sensor_CraneUp : BOOL := FALSE;
        Sensor_MagazinCapacitiveSensor : BOOL := FALSE;
        Sensor_MagazinEmergencyStop : BOOL := FALSE;
        Sensor_MagazinOpticalSensor : BOOL := FALSE;
        Sensor_MagazinSwitchManuellAutomatic : BOOL := FALSE;
        Sensor_SliderMovedOut : BOOL := FALSE;
        Sensor_SliderNotMovedOut : BOOL := FALSE;
        Sensor_StampEmergencyStop : BOOL := FALSE;
        Sensor_StampLowered : BOOL := FALSE;
        Sensor_StampSliderFilled : BOOL := FALSE;
        Sensor_StampSliderSensorMovedIn : BOOL := FALSE;
        Sensor_StampSliderSensorMovedOut : BOOL := FALSE;
        Sensor_StampStartButton : BOOL := FALSE;
        Sensor_StampSwitchManuellAutomatic : BOOL := FALSE;
        Sensor_StampUp : BOOL := FALSE;
        Sensor_StartButtonMagazin : BOOL := FALSE;
        Sensor_WorkpieceReady : BOOL := FALSE;
    END_VAR

    Mag.SliderNotMovedOut := Sensor_SliderNotMovedOut;
    Mag.SliderMovedOut := Sensor_SliderMovedOut;
    Mag.CraneOnMagazin := Sensor_CraneOnMagazin;
    Mag.CraneDown := Sensor_CraneDown;
    Mag.CraneUp := Sensor_CraneUp;
    Mag.CraneOnConveyor := Sensor_CraneOnConveyor;
    Mag.WorkpieceReady := Sensor_WorkpieceReady;
    Mag.StartButtonMagazin := Sensor_StartButtonMagazin;
    Actuator_MagazinSlider := Mag.MagazinSlider;
    Actuator_MagazinGreenLamp := Mag.MagazinGreenLamp;
    Crane.CraneUp := Sensor_CraneUp;
    Crane.CraneOnConveyor := Sensor_CraneOnConveyor;
    Crane.CraneDown := Sensor_CraneDown;
    Crane.CraneSucked := Sensor_CraneSucked;
    Crane.CraneOnMagazin := Sensor_CraneOnMagazin;
    Crane.MagazinCapacitiveSensor := Sensor_MagazinCapacitiveSensor;
    Crane.CranePositionStamp := Sensor_CranePositionStamp;
    Crane.SliderMovedOut := Sensor_SliderMovedOut;
    Crane.WorkpieceReady := Sensor_WorkpieceReady;
    Crane.MagazinOpticalSensor := Sensor_MagazinOpticalSensor;
    Crane.StampSliderFilled := Sensor_StampSliderFilled;
    Crane.StampSliderSensorMovedOut := Sensor_StampSliderSensorMovedOut;
    Crane.StampLowered := Sensor_StampLowered;
    Crane.StartButtonMagazin := Sensor_StartButtonMagazin;
    Actuator_CraneTurnCounterclockwise := Crane.CraneTurnCounterclockwise;
    Actuator_CraneTurnClockwise := Crane.CraneTurnClockwise;
    Actuator_CraneLower := Crane.CraneLower;
    Actuator_MagazinVacuumOff := Crane.MagazinVacuumOff;
    Actuator_MagazinVacuumOn := Crane.MagazinVacuumOn;
    Actuator_AnalogCranePressure := Crane.AnalogCranePressure;
    Stamp.StampSliderSensorMovedOut := Sensor_StampSliderSensorMovedOut;
    Stamp.StampSliderSensorMovedIn := Sensor_StampSliderSensorMovedIn;
    Stamp.StampSliderFilled := Sensor_StampSliderFilled;
    Stamp.StampUp := Sensor_StampUp;
    Stamp.StampLowered := Sensor_StampLowered;
    Stamp.CraneDown := Sensor_CraneDown;
    Stamp.CraneUp := Sensor_CraneUp;
    Stamp.CraneSucked := Sensor_CraneSucked;
    Stamp.CranePositionStamp := Sensor_CranePositionStamp;
    Stamp.CraneOnConveyor := Sensor_CraneOnConveyor;
    Stamp.StampStartButton := Sensor_StampStartButton;
    Actuator_StampSliderMovedOut := Stamp.StampSliderMovedOut;
    Actuator_StampSliderMovedIn := Stamp.StampSliderMovedIn;
    Actuator_StampWhiteLamp := Stamp.StampWhiteLamp;
    Actuator_StampPusher := Stamp.StampPusher;
    Actuator_StampGreenLamp := Stamp.StampGreenLamp;
    IF (Sensor_StampEmergencyStop AND Sensor_MagazinEmergencyStop) THEN
        Mag();
        Crane();
        Stamp();
        IF (Actuator_MagazinGreenLamp AND Actuator_StampGreenLamp) THEN
            IF ((Stamp.StartCommandStamp AND Crane.StartCommandCrane) AND Mag.StartCommandMagazin) THEN
                Crane.StartVar := TRUE;
                Mag.StartVar := TRUE;
                Stamp.StartVar := TRUE;
            END_IF
        END_IF
        Crane.SFCReset := FALSE;
        Mag.SFCReset := FALSE;
        Stamp.SFCReset := FALSE;
    ELSIF (NOT Sensor_StampEmergencyStop OR NOT Sensor_MagazinEmergencyStop) THEN
        Actuator_MagazinSlider := FALSE;
        Actuator_CraneLower := FALSE;
        Actuator_MagazinVacuumOn := FALSE;
        Actuator_MagazinVacuumOff := TRUE;
        Actuator_MagazinGreenLamp := FALSE;
        Actuator_CraneTurnCounterclockwise := FALSE;
        Actuator_CraneTurnClockwise := FALSE;
        Actuator_StampSliderMovedOut := TRUE;
        Actuator_StampSliderMovedIn := FALSE;
        Actuator_StampGreenLamp := FALSE;
        Actuator_StampPusher := FALSE;
        Actuator_AnalogCranePressure := INT#0;
        Crane.SFCReset := TRUE;
        Mag.SFCReset := TRUE;
        Stamp.SFCReset := TRUE;
        Crane.StartVar := FALSE;
        Mag.StartVar := FALSE;
        Stamp.StartVar := FALSE;
    END_IF
END_PROGRAM
FUNCTION_BLOCK CTD

    VAR_INPUT
        CD : BOOL := FALSE;
        LD : BOOL := FALSE;
        PV : INT := INT#0;
    END_VAR

    VAR_OUTPUT
        CV : INT := INT#0;
        Q : BOOL := FALSE;
    END_VAR

    IF LD THEN
        CV := PV;
    ELSIF (CU AND (CV > INT#0)) THEN
        CV := (CV - INT#1);
    END_IF
    Q := (CV <= INT#0);
END_FUNCTION_BLOCK

FUNCTION_BLOCK CTU

    VAR_INPUT
        CU : BOOL := FALSE;
        PV : INT := INT#0;
        R : BOOL := FALSE;
    END_VAR

    VAR_OUTPUT
        CV : INT := INT#0;
        Q : BOOL := FALSE;
    END_VAR

    IF R THEN
        CV := INT#0;
    ELSIF (CU AND (CV < PV)) THEN
        CV := (CV + INT#1);
    END_IF
    Q := (CV >= PV);
END_FUNCTION_BLOCK

FUNCTION_BLOCK R_TRIG

    VAR_INPUT
        CLK : BOOL := FALSE;
    END_VAR

    VAR
        M : BOOL := FALSE;
    END_VAR

    VAR_OUTPUT
        Q : BOOL := FALSE;
    END_VAR

    Q := (CLK AND NOT M);
    M := CLK;
END_FUNCTION_BLOCK

FUNCTION_BLOCK F_TRIG

    VAR_INPUT
        CLK : BOOL := FALSE;
    END_VAR

    VAR
        M : BOOL := TRUE;
    END_VAR

    VAR_OUTPUT
        Q : BOOL := FALSE;
    END_VAR

    Q := (NOT CLK AND NOT M);
    M := NOT CLK;
END_FUNCTION_BLOCK

FUNCTION SEL : ANY

    VAR_INPUT
        G : BOOL := FALSE;
        a : ANY;
        b : ANY;
    END_VAR

    VAR_OUTPUT
        SEL : ANY;
    END_VAR

    IF G THEN
        SEL := a;
    ELSE
        SEL := b;
    END_IF
END_FUNCTION

FUNCTION MAX : ANY_INT

    VAR_OUTPUT
        MAX : ANY_INT;
    END_VAR

    VAR_INPUT
        in0 : ANY_INT;
        in1 : ANY_INT;
    END_VAR

    MAX := sel((in0 >= in1), in0, in1);
END_FUNCTION

FUNCTION MIN : ANY_INT

    VAR_OUTPUT
        MIN : ANY_INT;
    END_VAR

    VAR_INPUT
        in0 : ANY_INT;
        in1 : ANY_INT;
    END_VAR

    MIN := sel((in0 <= in1), in0, in1);
END_FUNCTION

FUNCTION LIMIT : INT

    VAR_OUTPUT
        LIMIT : INT := INT#0;
    END_VAR

    VAR_INPUT
        in : ANY_INT;
        max : ANY_INT;
        min : ANY_INT;
    END_VAR

    LIMIT := MAX(min, MIN(in, max));
END_FUNCTION

FUNCTION ERROR : ANY

    VAR_OUTPUT
        ERROR : ANY;
    END_VAR

    VAR
        msg : STRING := WSTRING#"";
    END_VAR

END_FUNCTION

FUNCTION SMV : ANY

    VAR_OUTPUT
        SMV : ANY;
    END_VAR

    VAR_INPUT
        code : STRING := WSTRING#"";
    END_VAR

END_FUNCTION

FUNCTION_BLOCK TON

    VAR_OUTPUT
        ET : UINT := UINT#0;
        Q : BOOL := FALSE;
    END_VAR

    VAR_INPUT
        IN : BOOL := FALSE;
        PT : UINT := UINT#0;
    END_VAR

    IF IN THEN
        Q := (ET = UINT#0);
        IF (ET > UINT#0) THEN
            ET := (ET - UINT#1);
        ELSE
            ET := UINT#0;
        END_IF
    ELSE
        Q := FALSE;
        ET := PT;
    END_IF
END_FUNCTION_BLOCK

TYPE SFC_STEPS: STRUCT

        T :TIME
        X :BOOL
        _T :TIME
        _X :BOOLEND_STRUCT;

END_TYPE

TYPE
    STATES_CRANE : (Init, Start_Crane, Crane_Init, Crane_Init_2, Interstep, Interstep_2, TimeDelay, Interstep_3, Turn_Right, Magazin_Stop, Crane_Lower, Step0, Crane_Lift_Magazin, Crane_Turn_Left_NOT_Metallic, Crane_On_Conveyor, Stamp_Pressure_Profile_Set_Metallic, Crane_Lift_Magazin_Metallic, Crane_Turn_Left_Metallic, Crane_On_Stamp_Metallic, release_Workpiece, Crane_Go_Up, Stamp_Pressure_Profile_Set_White, Crane_Lift_Magazine_White, Crane_Turn_Left_White, Crane_On_Stamp_White, release_Workpiece_White, Crane_Go_Up_White, Step3, Step2, pause, Turn_Right_Black, Magazin_Stop_Black, Crane_Lift_NOT_Metallic_Black, Crane_Turn_Left_NOT_Metallic_Black, Crane_On_Conveyor_Not_Metallica_Black, release_Black, Crane_Lift_Conveyor_Black, Crane_Turn_Left_Back_To_Stamp, Crane_On_Stamp_Stop_Black, Step4, Reset_interconnect, Lower_Crane, Suck_At_Stamp, Crane_Lift_At_Stamp, Crane_Turn_Left_From_Stamp, Crane_On_Conveyor_Metallic, release, Crane_Lift_Conveyor, No_Workpiece_ready, Crane_Turn_Left_Metallic2, Crane_On_Stamp_Metallic2, Interstep_4, Crane_On_Stamp_Metallic2_Lower, Suck_At_Stamp2, Crane_Lift_At_Stamp2, Crane_Turn_Right_From_Stamp, Crane_On_Conveyor_Metallic2, release2, Crane_Lift_Conveyor2, Turn_Right_Final, Magazin_Stop_Final);
    STATES_MAGAZIN : (Init, Start_Magazin, Green_Lamp, Magazin_Init, Magazin_Init_2, Interstep, convey, Step0, Slider_Move_Back, Step1);
    STATES_STAMP : (Init, Start_Stamp, Green_Lamp, Stamp_Init_1, Stamp_Init_2, Stamp_Init_3, Stamp_Init_4, Interstep, Interstep_2, Step0, StampSliderBack, StampProcess, Step1, StampSliderForward, Step2);
END_TYPE
